(* IEC 61131-3 sources: MotionTestBenchMaster/Logical/00_AID/Libraries/System_Libraries/AsEPL, 3 files *)

(* ---- AsEPL.typ ---- *)
(********************************************************************
 * COPYRIGHT -- Bernecker + Rainer
 ********************************************************************
 * Library: AsEPL
 * File: AsEPL.typ
 * Author: B+R
 ********************************************************************
 * Data types of library AsEPL
 ********************************************************************)

TYPE
	EPL_I_TYPE : STRUCT			(*internal use*)
		init	: UDINT ;
		hdl	: UDINT ;
		st	: UDINT ;
		errInfo	: UDINT ;
		size	: UDINT ;
		bus	: USINT ;
		sl	: USINT ;
		ss	: USINT ;
		if_	: USINT ;
		nd	: USINT ;
		tid	: UDINT ;
	END_STRUCT;
END_TYPE

(* ---- AsEPL.fun ---- *)
(********************************************************************
 * COPYRIGHT -- Bernecker + Rainer
 ********************************************************************
 * Library: AsEPL
 * File: AsEPL.fun
 * Author: B+R
 ********************************************************************
 * Functions and function blocks of library AsEPL
 ********************************************************************)

{REDUND_CONTEXT} {REDUND_UNREPLICABLE} FUNCTION_BLOCK EplSDORead					(*reads node's object entries when using an SDO transfer*)
	VAR_INPUT
		enable	:BOOL;						(*enables execution*)
		pDevice	:REFERENCE TO STRING[80];	(*device name given as a pointer, e.g., "SL<x>.SS<y>.IF<z>"*)
		node	:USINT;						(*address of the node to be read (1-127 or 0 for local OD)*)
		index	:UINT;						(*number of the index entry to be read*)
		subindex	:USINT;					(*number of the subindex entry to be read*)
		pData	:UDINT;						(*pointer to the buffer for read data*)
		datalen	:UDINT;						(*maximum length of the data to be read*)
	END_VAR

	VAR_OUTPUT
		status	:UINT;						(*execution status: ERR_OK, ERR_FUB_ENABLE_FALSE, 0xXXXX = see help*)
		errorinfo	:UDINT;					(*SDO Abort Code, e.g., EPL_ERR_SDO_PROTOCOL_TIMEOUT, EPL_ERR_SDO_COMMAND_ID_INVALID, ..*)
		readlen	:UDINT;						(*length of the entry read*)
	END_VAR

	VAR
		intern	:EPL_I_TYPE;				(*internal variable*)
	END_VAR
END_FUNCTION_BLOCK

{REDUND_CONTEXT} {REDUND_UNREPLICABLE} FUNCTION_BLOCK EplSDOWrite					(*writes a node's object entries when using an SDO transfer*)
	VAR_INPUT
		enable	:BOOL;						(*enables execution*)
		pDevice	:REFERENCE TO STRING[80];	(*device name given as a pointer, e.g., "SL<x>.SS<y>.IF<z>"*)
		node	:USINT;						(*address of the node to be written (1-255 or 0 for local OD)*)
		index	:UINT;						(*number of the index entry to be written*)
		subindex	:USINT;					(*number of the subindex entry to be written*)
		pData	:UDINT;						(*pointer to the data to be written*)
		datalen	:UDINT;						(*length of the data to be written*)
	END_VAR

	VAR_OUTPUT
		status	:UINT;						(*execution status: ERR_OK, ERR_FUB_ENABLE_FALSE, 0xXXXX = see help*)
		errorinfo	:UDINT;					(*SDO abort code, e.g., EPL_ERR_SDO_PROTOCOL_TIMEOUT, EPL_ERR_SDO_COMMAND_ID_INVALID, ..*)
	END_VAR

	VAR
		intern	:EPL_I_TYPE;				(*internal variable*)
	END_VAR
END_FUNCTION_BLOCK

{REDUND_CONTEXT} {REDUND_UNREPLICABLE} FUNCTION_BLOCK EplGetLocalNodeID			(*queries the local node address of the PLC*)
	VAR_INPUT
		enable	:BOOL;						(*enables execution*)
		pDevice	:REFERENCE TO STRING[80];	(*device name given as a pointer, e.g., "SL<x>.SS<y>.IF<z>"*)
	END_VAR

	VAR_OUTPUT
		status	:UINT;						(*execution status: ERR_OK, ERR_FUB_ENABLE_FALSE, 0xXXXX = see help*)
		nodeid	:USINT;						(*local node number of the PLC*)
	END_VAR
END_FUNCTION_BLOCK

{REDUND_CONTEXT} {REDUND_UNREPLICABLE} FUNCTION_BLOCK EplCreateObject				(*creates a object at the given index/subindex*)
	VAR_INPUT
		enable	:BOOL;						(*enables execution*)
		pDevice	:REFERENCE TO STRING[80];	(*device name given as a pointer, e.g., "SL<x>.SS<y>.IF<z>"*)
		index	:UINT;						(*index of object*)
		subindex:USINT;						(*subindex of object*)
		datalen	:UDINT;						(*length of the object in octets*)
	END_VAR

	VAR_OUTPUT
		status	:UINT;						(*execution status: ERR_OK, ERR_FUB_ENABLE_FALSE, 0xXXXX = see help*)
	END_VAR
END_FUNCTION_BLOCK

{REDUND_CONTEXT} {REDUND_UNREPLICABLE} FUNCTION_BLOCK EplDeleteObject				(*creates a object at the given index/subindex*)
	VAR_INPUT
		enable	:BOOL;						(*enables execution*)
		pDevice	:REFERENCE TO STRING[80];	(*device name given as a pointer, e.g., "SL<x>.SS<y>.IF<z>"*)
		index	:UINT;						(*index of object*)
		subindex:USINT;						(*subindex of object*)
	END_VAR

	VAR_OUTPUT
		status	:UINT;						(*execution status: ERR_OK, ERR_FUB_ENABLE_FALSE, 0xXXXX = see help*)
	END_VAR
END_FUNCTION_BLOCK

(* ---- AsEPL.var ---- *)
(********************************************************************
 * COPYRIGHT -- Bernecker + Rainer
 ********************************************************************
 * Library: AsEPL
 * File: AsEPL.var
 * Author: B+R
 ********************************************************************
 * Local variables of library AsEPL
 ********************************************************************)

VAR CONSTANT
	ERR_ASEPL_BASE	: UINT	:= 31340;				(*base error number*)
	ERR_ASEPL_WRONG_DEVICE	: UINT	:= 31341;		(*specified device not a POWERLINK interface*)
	ERR_ASEPL_MN_ONLY	: UINT	:= 31342;			(*function can only be executed on an MN (managing node)*)
	ERR_ASEPL_CN_ONLY	: UINT	:= 31343;			(*function can only be executed on a CN (controlled node)*)
	ERR_ASEPL_ACCESS_FAILED	: UINT	:= 31344;		(*read or write access failed*)
	ERR_ASEPL_PARAM_OUTOFRANGE : UINT := 31345;		(*one or more parameters out of range*)
	ERR_ASEPL_INDEX_EXISTS : UINT := 31346;			(*index already exists*)
	ERR_ASEPL_SUBINDEX_EXISTS : UINT := 31347;		(*subindex already exists*)
	ERR_ASEPL_INDEX_DOESNOTEXIST : UINT := 31348;	(*index does not exist*)
	ERR_ASEPL_SUBINDEX_DOESNOTEXIST : UINT := 31349; (*subindex does not exists*)
	ERR_ASEPL_NILPOINTER : UINT := 31392;  (*nil pointer supplied*)
	ERR_ASEPL_NOT_IMPLEMENTED	: UINT	:= 31399; (*error code for non-implemented functionality*)
END_VAR
